Fanuc KAREL source: kb00041.compact.KL

PROGRAM KB00041
%STACKSIZE=65535
%PRIORITY=65535
%NOLOCKGROUP
VAR
P1 : STRING[80]
P2 : REAL
BEGIN
P1='A'
P2=1.0
CNV_STR_REAL(P1,P2)
END KB00041
